FUNCTION_BLOCK FB_LintBase
VAR_INPUT
END_VAR
VAR_OUTPUT
END_VAR
VAR
END_VAR

END_FUNCTION_BLOCK

(* stored: Version 1.1.0.1, ProductVersion 3.1.4026.18
   POU FB_LintBase: Id {90f3b172-1a65-092d-090e-17a5cb4bc037}, SpecialFunc None *)
